# EPICS substitutions: db/MicroEpsilon/ecmcOptoILD2300_100mm.substitutions
file "ecmc_analogInput-chX.template"
{
  pattern { CH_ID,  KEY,   EGU,  PREC,  ESLO, suffix    }
          { 01,     "Enc", "mm", 5,     1e-6, "-PosAct"  }
}
